(* IEC 61131-3 sources: llm-plc-st-eval/data/processed_definitivo/gemini-3.1-pro-preview/B2/zero_shot, 3 files *)

(* ---- ejec_1.st ---- *)
FUNCTION_BLOCK FB_Valvula
VAR_INPUT
    nivelAlto : BOOL; // Sensor de nivel alto del tanque
END_VAR
VAR_OUTPUT
    valvula : BOOL; // Comando para abrir (TRUE) o cerrar (FALSE) la válvula
END_VAR
VAR
    temporizador : TON; // Temporizador de retardo a la conexión (Timer On Delay)
END_VAR

// El temporizador se activa con el sensor de nivel alto.
// Si nivelAlto es TRUE por 5 segundos continuos, la salida Q del temporizador será TRUE.
// Si nivelAlto pasa a FALSE, el temporizador se reinicia y Q pasa a FALSE inmediatamente.
temporizador(IN := nivelAlto, PT := T#5S);

// La válvula se abre solo cuando el temporizador ha cumplido el tiempo establecido.
valvula := temporizador.Q;

END_FUNCTION_BLOCK

(* ---- ejec_2.st ---- *)
FUNCTION_BLOCK FB_Valvula
VAR_INPUT
    nivelAlto : BOOL; // Indica si el sensor de nivel alto está activo
END_VAR

VAR_OUTPUT
    valvula : BOOL; // Comando para abrir (TRUE) o cerrar (FALSE) la válvula de drenaje
END_VAR

VAR
    temporizador : TON; // Temporizador con retardo a la conexión (On-Delay)
END_VAR

// El temporizador evalúa si el nivel alto se mantiene activo por 5 segundos continuos.
// Si nivelAlto pasa a FALSE, el temporizador se reinicia y su salida Q pasa a FALSE de inmediato.
temporizador(IN := nivelAlto, PT := T#5S);

// La válvula se abre solo cuando el temporizador ha cumplido el tiempo establecido.
valvula := temporizador.Q;

END_FUNCTION_BLOCK

(* ---- ejec_3.st ---- *)
FUNCTION_BLOCK FB_Valvula
VAR_INPUT
    nivelAlto : BOOL; // Señal del sensor de nivel alto
END_VAR

VAR_OUTPUT
    valvula : BOOL;   // Comando para abrir (TRUE) o cerrar (FALSE) la válvula
END_VAR

VAR
    tonRetardo : TON; // Temporizador de retardo a la conexión (Timer On Delay)
END_VAR

// Configuración y ejecución del temporizador
// IN: Inicia el conteo si nivelAlto es TRUE. Se resetea inmediatamente si es FALSE.
// PT: Tiempo de retardo establecido en 5 segundos.
tonRetardo(IN := nivelAlto, PT := T#5S);

// La salida del temporizador (Q) se activa tras 5 segundos continuos de nivel alto.
// Si nivelAlto pasa a FALSE, Q se desactiva de inmediato, cerrando la válvula.
valvula := tonRetardo.Q;

END_FUNCTION_BLOCK
